(* IEC 61131-3 sources: axsharp/src/AXSharp.compiler/tests/AXSharp.Compiler.CsTests/samples/units/src, 39 files *)

(* ---- compileromitsattribute.st ---- *)
NAMESPACE CompilerOmmits
    {S7.extern=ReadWrite}
    CLASS ClassWithArrays
        VAR PUBLIC
            {#ix-attr:[CompilerOmitsAttribute()]}
            _must_be_omitted_everywhere : Complex;
            {#ix-attr:[CompilerOmitsAttribute("Onliner")]}
            _must_be_omitted_in_onliner : Complex;
            {#ix-attr:[CompilerOmitsAttribute("POCO")]}
             _must_be_omitted_in_poco : Complex;
            _primitive  : ARRAY[0..10] OF BYTE;
        END_VAR

    END_CLASS

    {S7.extern=ReadWrite}
    CLASS PUBLIC Complex
        VAR PUBLIC
            HelloString : STRING;
            Id : ULINT;
        END_VAR
    END_CLASS
END_NAMESPACE

NAMESPACE CompilerOmmitsEnums
    {S7.extern=ReadWrite}
    CLASS ClassWithEnums
        VAR PUBLIC
            colors : Colors;
            NamedValuesColors : NamedValuesColors;
        END_VAR

    END_CLASS

    TYPE
        Colors : (Red, Green, Blue) := Red;
    END_TYPE

    TYPE
        NamedValuesColors : STRING (Red := '1', Green := '2', Blue := '3') := Red;
    END_TYPE

END_NAMESPACE

NAMESPACE CompilerOmmitsMisc
    {S7.extern=ReadWrite}
    CLASS PUBLIC VariousMembers
        VAR PUBLIC
            _SomeClass : SomeClass;
            _Motor : ComersMotor;
        END_VAR
    END_CLASS

    {S7.extern=ReadWrite}
    CLASS SomeClass
        VAR PUBLIC
            SomeClassVariable : STRING;
        END_VAR
    END_CLASS

    TYPE
        {S7.extern=ReadWrite}
        ComersMotor : STRUCT
            isRunning : BOOL;
        END_STRUCT;
        {S7.extern=ReadWrite}
        ComersVehicle : STRUCT
            m : ComersMotor;
            displacement : INT;
        END_STRUCT;
    END_TYPE
END_NAMESPACE

NAMESPACE CompilerOmmitsUnknownArrays
    {S7.extern=ReadWrite}
    CLASS ClassWithArrays
        VAR PUBLIC
            _complexKnown : ARRAY[0..10] OF Complex;
            _complexUnknown : ARRAY [0..10] OF ComplexUnknown;
            _primitive  : ARRAY[0..10] OF BYTE;
        END_VAR

    END_CLASS

    {S7.extern=ReadWrite}
    CLASS PUBLIC Complex
        VAR PUBLIC
            HelloString : STRING;
            Id : ULINT;
        END_VAR
    END_CLASS
END_NAMESPACE

(* ---- enum_simple.st ---- *)
TYPE
    Colors : (Red, Green, Blue) := Red;
END_TYPE

(* ---- misc.st ---- *)
NAMESPACE Enums
{S7.extern=ReadWrite}
    CLASS ClassWithEnums
        VAR PUBLIC
            colors : Colors;
            NamedValuesColors : NamedValuesColors;
        END_VAR

    END_CLASS

    TYPE
        Colors : (Red, Green, Blue) := Red;
    END_TYPE

    TYPE
        NamedValuesColors : STRING (Red := '1', Green := '2', Blue := '3') := Red;
    END_TYPE

END_NAMESPACE

NAMESPACE misc
{S7.extern=ReadWrite}
    CLASS PUBLIC VariousMembers
        VAR PUBLIC
            _SomeClass : SomeClass;
            _Motor : MiscMotor;
        END_VAR
    END_CLASS

    {S7.extern=ReadWrite}
    CLASS SomeClass
        VAR PUBLIC
            SomeClassVariable : STRING;
        END_VAR
    END_CLASS

    TYPE
        {S7.extern=ReadWrite}
        MiscMotor : STRUCT
            isRunning : BOOL;
        END_STRUCT;
        {S7.extern=ReadWrite}
        MiscVehicle : STRUCT
            m : MiscMotor;
            displacement : INT;
        END_STRUCT;
    END_TYPE
END_NAMESPACE

NAMESPACE UnknownArraysShouldNotBeTraspiled
    {S7.extern=ReadWrite}
    CLASS ClassWithArrays
        VAR PUBLIC
            _complexKnown : ARRAY[0..10] OF Complex;
            _complexUnknown : ARRAY [0..10] OF ComplexUnknown;
            _primitive  : ARRAY[0..10] OF BYTE;
        END_VAR

    END_CLASS

    {S7.extern=ReadWrite}
    CLASS PUBLIC Complex
        VAR PUBLIC
            HelloString : STRING;
            Id : ULINT;
        END_VAR
    END_CLASS
END_NAMESPACE

(* ---- mixed_access.st ---- *)
CONFIGURATION config
    VAR_GLOBAL
        {S7.extern=ReadWrite}
        MotorOn : BOOL;             // variable can be read and written

        {S7.extern=ReadOnly}
        MotorState: INT;            // variable can only be read

        MotorFlags: UINT;           // variable is not accessible by an external system (default: hidden)

        {S7.extern=ReadWrite}
        Motor1 : MixedAccessMotor;        // the variables in Motor1 be read and written if enabled

        {S7.extern=ReadOnly}
        Motor2 : MixedAccessMotor;        // the variables in Motor2 be only read if enabled

        {S7.extern=ReadWrite}
        s1 : struct1;
        {S7.extern=ReadWrite}
        s4 : struct4;

        {S7.extern=ReadWrite}
        mot1 : SpecificMotorA;
    END_VAR
END_CONFIGURATION

CLASS MixedAccessMotor
    VAR PUBLIC
        {S7.extern=ReadWrite}
        Run               : BOOL;
        ReverseDirection  : BOOL;
    END_VAR
    VAR INTERNAL
        {S7.extern=ReadOnly}
        ActualVelocity    : LReal;
    END_VAR
    // ...
END_CLASS

TYPE
    struct1 : STRUCT  {S7.extern=ReadWrite}  s2 : struct2;   END_STRUCT;
    struct2 : STRUCT  {S7.extern=ReadOnly}   s3 : struct3;   END_STRUCT;
    struct3 : STRUCT  {S7.extern=ReadWrite}  s4 : struct4;   END_STRUCT;
    struct4 : STRUCT  {S7.extern=ReadWrite}  s5 : INT;       END_STRUCT;
END_TYPE

{S7.extern=ReadWrite}
CLASS ABSTRACT AbstractMotor
    VAR PUBLIC
        Run               : BOOL;
        ReverseDirection  : BOOL;
    END_VAR
    ...
END_CLASS

{S7.extern=ReadWrite}
CLASS GenericMotor  EXTENDS AbstractMotor
    VAR INTERNAL
        {S7.extern=ReadOnly}
        ActualVelocity    : LReal;
    END_VAR
    ...
END_CLASS

{S7.extern=ReadWrite}
CLASS SpecificMotorA  EXTENDS GenericMotor
    VAR INTERNAL
        {S7.extern=ReadWrite}
        MaxAcceleration    : LReal;
    END_VAR
    ...
END_CLASS

(* ---- struct_simple.st ---- *)
TYPE
    {S7.extern=ReadWrite}
    StructSimpleMotor : STRUCT
        isRunning : BOOL;
    END_STRUCT;
    {S7.extern=ReadWrite}
    StructSimpleVehicle : STRUCT
        m : StructSimpleMotor;
        displacement : INT;
    END_STRUCT;
END_TYPE

(* ---- type_named_values.st ---- *)
NAMESPACE NamedValuesNamespace
    TYPE
        LightColors : INT (
            LRED := 12,
            LGREEN := 14,
            LBLUE := 23
        );
    END_TYPE

    {S7.extern=ReadWrite}
    CLASS PUBLIC using_type_named_values
        VAR PUBLIC
            LColors : LightColors;
        END_VAR
    END_CLASS
END_NAMESPACE

(* ---- type_named_values_literals.st ---- *)
NAMESPACE Simatic.Ax.StateFramework
    TYPE
        StateControllerStatus : WORD (
            STATUS_NO_ERR := WORD#16#7000,
            STATUS_IS_RUNNING := WORD#16#7001,
            STATUS_STATE_CHANGED := WORD#16#7002,
            STATUS_NO_INITIALSTATE := WORD#16#8100,
            STATUS_NO_NEXTSTATE := WORD#16#8101
        ) := STATUS_NO_ERR;
    END_TYPE

    {S7.extern=ReadWrite}
    CLASS PUBLIC using_type_named_values
        VAR PUBLIC
            LColors : StateControllerStatus;
        END_VAR
    END_CLASS
END_NAMESPACE

(* ---- type_with_enum.st ---- *)
NAMESPACE Simatic.Ax.StateFramework
    INTERFACE IGuard

        METHOD Check : BOOL
        END_METHOD

        METHOD Reset
        END_METHOD

    END_INTERFACE
END_NAMESPACE

NAMESPACE Simatic.Ax.StateFramework

    /// Condition
    /// GT: Greater than compareValue
    /// EQ: Equal to compareValue
    /// LT: Less than compareValue
    /// NE: Is not equal to compareValue
    /// GE: Greater or equal to compareValue
    /// LE: Less or equal to compareValue
    TYPE
        Condition : (GT, EQ, LT, NE, GE, LE);
    END_TYPE

    {S7.extern=ReadWrite}
    CLASS CompareGuardLint IMPLEMENTS IGuard
        VAR PUBLIC
            Value : REF_TO LINT;
            CompareToValue : LINT;
            Condition : Condition;
        END_VAR

        METHOD PUBLIC Config
            VAR_INPUT
                countValue : REF_TO LINT;
                compareValue : LINT;
                compareCondition : Condition;
            END_VAR
            Value := countValue;
            CompareToValue := compareValue;
            Condition := compareCondition;
        END_METHOD

        // ---------------- IMPLEMENT IGuard---------------------------
        METHOD PUBLIC Check : BOOL

            CASE Condition OF
                Condition#GT : Check := Value^ > CompareToValue;
                Condition#EQ : Check := Value^ = CompareToValue;
                Condition#LT : Check := Value^ < CompareToValue;
                Condition#GE : Check := Value^ >= CompareToValue;
                Condition#LE : Check := Value^ <= CompareToValue;
            END_CASE
            ;

        END_METHOD

        METHOD PUBLIC Reset
            ;
        END_METHOD
        // ---------------- END IMPLEMENT IGuard---------------------------

    END_CLASS
END_NAMESPACE

(* ---- types_with_name_attributes.st ---- *)
NAMESPACE TypeWithNameAttributes
    TYPE
        {#ix-attr:[Container(Layout.Wrap)]}
        {S7.extern=ReadWrite}
        TypesNameAttrMotor : STRUCT
            isRunning : BOOL;
        END_STRUCT;
        {S7.extern=ReadWrite}
        TypesNameAttrVehicle : STRUCT
            m : TypesNameAttrMotor;
            displacement : INT;
        END_STRUCT;
    END_TYPE

    {#ix-prop:public string AttributeName}
    {S7.extern=ReadWrite}
    CLASS NoAccessModifierClass
        VAR PUBLIC
            SomeClassVariable : STRING;
        END_VAR
    END_CLASS
END_NAMESPACE

(* ---- class_extends_and_implements.st ---- *)
{S7.extern=ReadWrite}
CLASS PUBLIC ExtendsAndImplements EXTENDS ExtendeeExtendsAndImplements IMPLEMENTS IImplementation1, IImplementation2

END_CLASS

{S7.extern=ReadWrite}
CLASS PUBLIC ExtendeeExtendsAndImplements

END_CLASS

INTERFACE PUBLIC IImplementation1 END_INTERFACE
INTERFACE PUBLIC IImplementation2 END_INTERFACE

(* ---- class_implements.st ---- *)
{S7.extern=ReadWrite}
CLASS PUBLIC _NULL_CONTEXT IMPLEMENTS IContext

END_CLASS

INTERFACE PUBLIC IContext

END_INTERFACE

(* ---- class_implements_multiple.st ---- *)
{S7.extern=ReadWrite}
CLASS PUBLIC _NULL_CONTEXT_MULTIPLE IMPLEMENTS IContext_Multiple, IObject_Multiple

END_CLASS

INTERFACE PUBLIC IContext_Multiple

END_INTERFACE

INTERFACE PUBLIC IObject_Multiple

END_INTERFACE

(* ---- file_with_unsupported.st ---- *)
NAMESPACE Unsupported
  FUNCTION SomeFunction : INT
    ;
  END_FUNCTION
END_NAMESPACE

(* ---- abstract_members.st ---- *)
{S7.extern=ReadWrite}
CLASS ABSTRACT AbstractMembersMotor
    VAR PUBLIC
        Run               : BOOL;
        ReverseDirection  : BOOL;
    END_VAR
    ...
END_CLASS

(* ---- array_declaration.st ---- *)
NAMESPACE ArrayDeclarationSimpleNamespace
    {S7.extern=ReadWrite}
    CLASS array_declaration_class
        VAR PUBLIC
            primitive : ARRAY[1..100] OF INT;
            complex : ARRAY[1..100] OF some_complex_type;
            // multidimensional arrays should not be transpiled
            complex_multidim : ARRAY[1..100, 0..30] OF some_complex_type;
            primitive_multidim : ARRAY[1..100, 0..100, 0..300] OF INT;
        END_VAR
    END_CLASS
    {S7.extern=ReadWrite}
    CLASS some_complex_type
        VAR

        END_VAR

    END_CLASS

END_NAMESPACE

(* ---- class_all_primitives.st ---- *)
{S7.extern=ReadWrite}
CLASS class_all_primitives
    VAR PUBLIC
        myBOOL	        :       BOOL	      ;
        myBYTE	        :       BYTE	      ;
        myWORD	        :       WORD	      ;
        myDWORD	        :       DWORD	      ;
        myLWORD	        :       LWORD	      ;
        mySINT	        :       SINT	      ;
        myINT	        :       INT	          ;
        myDINT	        :       DINT	      ;
        myLINT	        :       LINT	      ;
        myUSINT	        :       USINT	      ;
        myUINT	        :       UINT	      ;
        myUDINT	        :       UDINT	      ;
        myULINT	        :       ULINT	      ;
        myREAL	        :       REAL	      ;
        myLREAL	        :       LREAL	      ;
        myTIME	        :       TIME	      ;
        myLTIME	        :       LTIME	      ;
        myDATE	        :       DATE	      ;
     //   myLDATE	        :       LDATE	      ;
        myTIME_OF_DAY	:       TIME_OF_DAY	  ;
     //   myLTIME_OF_DAY	:       LTIME_OF_DAY  ;
        myDATE_AND_TIME  :      DATE_AND_TIME ;
     //   myLDATE_AND_TIME :      LDATE_AND_TIME;
     //   myCHAR	        :       CHAR	      ;
     //   myWCHAR	        :       WCHAR	      ;
        mySTRING	        :   STRING	      ;
        myWSTRING	    :       WSTRING	      ;
    END_VAR
END_CLASS

(* ---- class_extended_by_known_type.st ---- *)
USING Simatic.Ax.Stateframework;
USING Simatic.Ax.StatePattern;

NAMESPACE Simatic.Ax.StateFramework
    {S7.extern=ReadWrite}
    CLASS State1Transition EXTENDS AbstractState

        METHOD PUBLIC OVERRIDE OnEntry
            ;
        END_METHOD

        METHOD PUBLIC OVERRIDE OnExit
            ;
        END_METHOD

        METHOD PUBLIC OVERRIDE Action
            ;
        END_METHOD

    END_CLASS

END_NAMESPACE

NAMESPACE Simatic.Ax.StateFramework
    {S7.extern=ReadWrite}
    CLASS ABSTRACT AbstractState IMPLEMENTS IState, IStateMuteable

        VAR PUBLIC
            Transition1 : ITransition;
            StateID : INT;
            StateName : String;
        END_VAR

        VAR PROTECTED
             _actualStatus : StateStatus;
        END_VAR

        // METHOD PUBLIC ABSTRACT OnEntry
        // END_METHOD
        METHOD PUBLIC OnEntry
            _actualStatus := StateStatus#Active;
        END_METHOD

        METHOD PUBLIC ABSTRACT OnExit
        END_METHOD

        METHOD PUBLIC ABSTRACT Action
        END_METHOD

        METHOD PUBLIC GetTransition : ITransition
            VAR_INPUT
                pos : UINT;
            END_VAR
            IF (THIS.TransitionCount() = pos + UINT#1) THEN
                GetTransition := transition1;
            ELSE
                GetTransition := NULL;
            END_IF;
        END_METHOD

        METHOD PUBLIC TransitionCount : UINT
            IF (transition1 <> NULL) THEN
                TransitionCount := UINT#1;
            ELSE
                TransitionCount := UINT#0;
            END_IF;
        END_METHOD

        METHOD PUBLIC GetStateID : INT
            GetStateID := StateID;
        END_METHOD

        METHOD PUBLIC FINAL GetStateName : STRING
            GetStateName := StateName;
        END_METHOD

        METHOD PUBLIC FINAL GetStatus : StateStatus
            GetStatus := _actualStatus;
        END_METHOD

        METHOD PUBLIC FINAL SetStatus
            VAR_INPUT
                status : StateStatus;
            END_VAR
            _actualStatus := status;
        END_METHOD
    END_CLASS
END_NAMESPACE

(* ---- class_extends.st ---- *)
{S7.extern=ReadWrite}
CLASS PUBLIC Extended EXTENDS Extendee

END_CLASS

{S7.extern=ReadWrite}
CLASS PUBLIC Extendee

END_CLASS

(* ---- class_generic_extension.st ---- *)
NAMESPACE Generics
    {#ix-generic:<TOnline, TPlain> where TOnline : ITwinObject}
    {S7.extern=ReadWrite}
    CLASS PUBLIC Extender

    END_CLASS

    {S7.extern=ReadWrite}
    CLASS PUBLIC Extendee EXTENDS Extender
        VAR PUBLIC
            {#ix-generic:TOnline}
            SomeType : SomeType;
            {#ix-generic:TPlain as POCO}
            SomeTypeAsPoco : SomeType;
        END_VAR
    END_CLASS

    {S7.extern=ReadWrite}
    CLASS PUBLIC Extendee2 EXTENDS Extender
        VAR PUBLIC
            {#ix-generic:TOnline}
            {#ix-generic:TPlain as POCO}
            SomeType : SomeType;
        END_VAR
    END_CLASS

    {S7.extern=ReadWrite}
    CLASS SomeType
    END_IF;
END_NAMESPACE

(* ---- class_internal.st ---- *)
{S7.extern=ReadWrite}
CLASS INTERNAL ClassWithComplexTypes

END_CLASS

(* ---- class_no_access_modifier.st ---- *)
{S7.extern=ReadWrite}
CLASS NoAccessModifierClass

END_CLASS

(* ---- class_with_complex_members.st ---- *)
NAMESPACE ClassWithComplexTypesNamespace
    {S7.extern=ReadWrite}
    CLASS PUBLIC ClassWithComplexTypes
        VAR PUBLIC
           myComplexType : ComplexType1;
        END_VAR
    END_CLASS

    {S7.extern=ReadWrite}
    CLASS PUBLIC ComplexType1

    END_CLASS
END_NAMESPACE

(* ---- class_with_constant_members.st ---- *)
NAMESPACE ClassWithConstantMembersNamespace
    {S7.extern=ReadWrite}
    CLASS PUBLIC ClassWithConstantMembers
        VAR PUBLIC
           myNonConstant : INT;
        END_VAR
        VAR CONSTANT
           myConstant : INT := 10;
           myConstantString : STRING := 'hello';
        END_VAR
    END_CLASS
END_NAMESPACE

(* ---- class_with_non_public_members.st ---- *)
NAMESPACE ClassWithNonTraspilableMemberssNamespace
   {S7.extern=ReadWrite}
    CLASS PUBLIC ClassWithNonTraspilableMembers
        VAR PUBLIC
           myComplexType : ComplexType1;
        END_VAR

        VAR
           myComplexType1 : ComplexType1;
           myBooool : BOOL;
        END_VAR

        VAR
           myComplexType2 : ComplexType1;
           myBooool1 : BOOL;
        END_VAR
    END_CLASS
    {S7.extern=ReadWrite}
    CLASS PUBLIC ComplexType1

    END_CLASS
END_NAMESPACE

(* ---- class_with_pragmas.st ---- *)
NAMESPACE ClassWithPragmasNamespace
    {#ix-attr:[Container(Layout.Stack)]}
    {S7.extern=ReadWrite}
    CLASS PUBLIC  ClassWithPragmas
        VAR PUBLIC
           {#ix-attr:[Container(Layout.Wrap)]}
           {S7.extern=ReadWrite}
           myComplexType : ComplexType1;
        END_VAR
    END_CLASS

    CLASS PUBLIC ComplexType1

    END_CLASS
END_NAMESPACE

(* ---- class_with_primitive_members.st ---- *)
NAMESPACE ClassWithPrimitiveTypesNamespace
    {S7.extern=ReadWrite}
    CLASS PUBLIC ClassWithPrimitiveTypes
        VAR PUBLIC
           myBOOL	        :       BOOL	      ;
           myBYTE	        :       BYTE	      ;
           myWORD	        :       WORD	      ;
           myDWORD	        :       DWORD	      ;
           myLWORD	        :       LWORD	      ;
           mySINT	        :       SINT	      ;
           myINT	        :       INT	          ;
           myDINT	        :       DINT	      ;
           myLINT	        :       LINT	      ;
           myUSINT	        :       USINT	      ;
           myUINT	        :       UINT	      ;
           myUDINT	        :       UDINT	      ;
           myULINT	        :       ULINT	      ;
           myREAL	        :       REAL	      ;
           myLREAL	        :       LREAL	      ;
           myTIME	        :       TIME	      ;
           myLTIME	        :       LTIME	      ;
           myDATE	        :       DATE	      ;
           myLDATE	        :       LDATE	      ;
           myTIME_OF_DAY	:       TIME_OF_DAY	  ;
           myLTIME_OF_DAY	:       LTIME_OF_DAY  ;
           myDATE_AND_TIME  :       DATE_AND_TIME ;
           myLDATE_AND_TIME :       LDATE_AND_TIME;
           myCHAR	        :       CHAR	      ;
           myWCHAR	        :       WCHAR	      ;
           mySTRING	        :       STRING	      ;
           myWSTRING	    :       WSTRING	      ;
        END_VAR
    END_CLASS
END_NAMESPACE

(* ---- class_with_using_directives.st ---- *)
{S7.extern=ReadWrite}
CLASS INTERNAL ClassWithUsingDirectives
    USING SimpleFirstLevelNamespace, SimpleQualifiedNamespace.Qualified;
    USING HelloLevelOne.HelloLevelTwo;
    USING InexistingNamespace;
END_CLASS

NAMESPACE SimpleFirstLevelNamespace

END_NAMESPACE

NAMESPACE SimpleQualifiedNamespace.Qualified

END_NAMESPACE

NAMESPACE HelloLevelOne
    NAMESPACE HelloLevelTwo
    END_NAMESPACE
END_NAMESPACE

(* ---- configuration.st ---- *)
CONFIGURATION MyConfiguration
    TASK Main(Interval := T#1000ms, Priority := 1);
    PROGRAM P1 WITH Main: MyProgram;

    VAR_GLOBAL
        {S7.extern=ReadWrite}
        Complex : ComplexForConfig;
        {S7.extern=ReadWrite}
        myBOOL	        :       BOOL	      ;
        {S7.extern=ReadWrite}
        myBYTE	        :       BYTE	      ;
        {S7.extern=ReadWrite}
        myWORD	        :       WORD	      ;
        {S7.extern=ReadWrite}
        myDWORD	        :       DWORD	      ;
        {S7.extern=ReadWrite}
        myLWORD	        :       LWORD	      ;
        {S7.extern=ReadWrite}
        mySINT	        :       SINT	      ;
        {S7.extern=ReadWrite}
        myINT	        :       INT	          ;
        {S7.extern=ReadWrite}
        myDINT	        :       DINT	      ;
        {S7.extern=ReadWrite}
        myLINT	        :       LINT	      ;
        {S7.extern=ReadWrite}
        myUSINT	        :       USINT	      ;
        {S7.extern=ReadWrite}
        myUINT	        :       UINT	      ;
        {S7.extern=ReadWrite}
        myUDINT	        :       UDINT	      ;
        {S7.extern=ReadWrite}
        myULINT	        :       ULINT	      ;
        {S7.extern=ReadWrite}
        myREAL	        :       REAL	      ;
        {S7.extern=ReadWrite}
        myLREAL	        :       LREAL	      ;
        {S7.extern=ReadWrite}
        myTIME	        :       TIME	      ;
        {S7.extern=ReadWrite}
        myLTIME	        :       LTIME	      ;
        {S7.extern=ReadWrite}
        myDATE	        :       DATE	      ;
        {S7.extern=ReadWrite}
        myLDATE	        :       LDATE	      ;
        {S7.extern=ReadWrite}
        myTIME_OF_DAY	:       TIME_OF_DAY	  ;
        {S7.extern=ReadWrite}
        myLTIME_OF_DAY	:       LTIME_OF_DAY  ;
        {S7.extern=ReadWrite}
        myDATE_AND_TIME  :       DATE_AND_TIME ;
        {S7.extern=ReadWrite}
        myLDATE_AND_TIME :       LDATE_AND_TIME;
        {S7.extern=ReadWrite}
        myCHAR	        :       CHAR	      ;
        {S7.extern=ReadWrite}
        myWCHAR	        :       WCHAR	      ;
        {S7.extern=ReadWrite}
        mySTRING	        :       STRING	      ;
        {S7.extern=ReadWrite}
        myWSTRING	    :       WSTRING	      ;
        {S7.extern=ReadWrite}
        mySTRING_10	    :       STRING[10]	  ;
        {S7.extern=ReadWrite}
        myWSTRING_10	:       WSTRING[10]	  ;

        {S7.extern=ReadWrite}
        {#ix-attr:[ReadOnce()]}
        myWSTRING_readOnce	    :       WSTRING	      ;
        {#ix-attr:[ReadOnly()]}
        {S7.extern=ReadWrite}
        myWSTRING_readOnly	    :       WSTRING	      ;
        {#ix-attr:[ReadOnce()]}
        {S7.extern=ReadWrite}
        cReadOnce           : ComplexForConfig;
        {#ix-attr:[ReadOnly()]}
        {S7.extern=ReadWrite}
        cReadOnly           : ComplexForConfig;
        {S7.extern=ReadWrite}
        Colorss : Colorss;
        {S7.extern=ReadWrite}
        Colorsss : Colorsss;

        {S7.extern=ReadWrite}
        {#ix-attr:[CompilerOmitsAttribute()]}
        _must_be_omitted_everywhere : BOOL;
        {S7.extern=ReadWrite}
        {#ix-attr:[CompilerOmitsAttribute("Onliner")]}
        _must_be_omitted_in_onliner : BOOL;
        {S7.extern=ReadWrite}
        {#ix-attr:[CompilerOmitsAttribute("POCO")]}
         _must_be_omitted_in_poco : BOOL;
    END_VAR
END_CONFIGURATION

CONFIGURATION MyConfiguration2
    VAR_GLOBAL
        {S7.extern=ReadWrite}
        Colorss2 : Colorss;
        {S7.extern=ReadWrite}
        Colorsss2 : Colorsss;
    END_VAR
END_CONFIGURATION

{S7.extern=ReadWrite}
CLASS PUBLIC ComplexForConfig
    VAR PUBLIC
        myBOOL	        :       BOOL	      ;
        myBYTE	        :       BYTE	      ;
        myWORD	        :       WORD	      ;
        myDWORD	        :       DWORD	      ;
        myLWORD	        :       LWORD	      ;
        mySINT	        :       SINT	      ;
        myINT	        :       INT	          ;
        myDINT	        :       DINT	      ;
        myLINT	        :       LINT	      ;
        myUSINT	        :       USINT	      ;
        myUINT	        :       UINT	      ;
        myUDINT	        :       UDINT	      ;
        myULINT	        :       ULINT	      ;
        myREAL	        :       REAL	      ;
        myLREAL	        :       LREAL	      ;
        myTIME	        :       TIME	      ;
        myLTIME	        :       LTIME	      ;
        myDATE	        :       DATE	      ;
        myLDATE	        :       LDATE	      ;
        myTIME_OF_DAY	:       TIME_OF_DAY	  ;
        myLTIME_OF_DAY	:       LTIME_OF_DAY  ;
        myDATE_AND_TIME  :       DATE_AND_TIME ;
        myLDATE_AND_TIME :       LDATE_AND_TIME;
        myCHAR	        :       CHAR	      ;
        myWCHAR	        :       WCHAR	      ;
        mySTRING	        :       STRING	      ;
        myWSTRING	    :       WSTRING	      ;
        myMotor         : ConfigMotor;
    END_VAR
END_CLASS

TYPE
    Colorss : (Red, Green, Blue) := Red;
END_TYPE

TYPE
    Colorsss : ULINT (Red := ULINT#1, Green := ULINT#2, Blue := ULINT#3) := Red;
END_TYPE

 TYPE
        {S7.extern=ReadWrite}
        ConfigMotor : STRUCT
            isRunning : BOOL;
        END_STRUCT;
        {S7.extern=ReadWrite}
        ConfigVehicle : STRUCT
            m : ConfigMotor;
            displacement : INT;
        END_STRUCT;
    END_TYPE

(* ---- file_with_usings.st ---- *)
USING FileWithUsingsSimpleFirstLevelNamespace;
USING FileWithUsingsSimpleQualifiedNamespace.Qualified;
USING FileWithUsingsHelloLevelOne.FileWithUsingsHelloLevelTwo;

NAMESPACE FileWithUsingsSimpleFirstLevelNamespace
    CLASS Hello
        VAR

        END_VAR
    END_CLASS
END_NAMESPACE

NAMESPACE FileWithUsingsSimpleQualifiedNamespace.Qualified
    CLASS Hello
        VAR

        END_VAR
    END_CLASS
END_NAMESPACE

NAMESPACE FileWithUsingsHelloLevelOne
    NAMESPACE FileWithUsingsHelloLevelTwo
        CLASS Hello
            VAR

            END_VAR
        END_CLASS
    END_NAMESPACE
END_NAMESPACE

NAMESPACE ExampleNamespace
    CLASS Hello
        VAR
            a : FileWithUsingsSimpleFirstLevelNamespace.Hello;
            b : FileWithUsingsSimpleQualifiedNamespace.Qualified.Hello;
            c : FileWithUsingsHelloLevelOne.FileWithUsingsHelloLevelTwo.Hello;
        END_VAR
    END_CLASS
END_NAMESPACE

(* ---- generics.st ---- *)
// GENERIC
NAMESPACE GenericsTests
    {#ix-generic:<TOnline, TPlain> where TOnline : ITwinObject}
	{S7.extern=ReadWrite}
    CLASS PUBLIC Extender

    END_CLASS

    {S7.extern=ReadWrite}
	CLASS PUBLIC SomeTypeToBeGeneric
	     VAR PUBLIC
		    Boolean : BOOL;
			Cele : INT;
		 END_VAR
	END_CLASS

	{S7.extern=ReadWrite}
   CLASS PUBLIC Extendee2 EXTENDS Extender
        VAR PUBLIC
            {#ix-generic:TOnline}
            {#ix-generic:TPlain as POCO}
            {#ix-attr:[AXOpen.Data.AxoDataEntityAttribute]}
            {#ix-attr:[Container(Layout.Stack)]}
            {#ix-set:AttributeName = "Shared Header"}
            SomeData : SomeTypeToBeGeneric;
        END_VAR
   END_CLASS
END_NAMESPACE

(* ---- makereadonce.st ---- *)
NAMESPACE makereadonce
    {S7.extern=ReadWrite}
    CLASS PUBLIC MembersWithMakeReadOnce
        VAR PUBLIC
            {#ix-attr:[ReadOnce()]}
            makeReadOnceMember : STRING;
            someOtherMember : STRING;

            {#ix-attr:[ReadOnce()]}
            makeReadComplexMember : ComplexMember;
            someotherComplexMember : ComplexMember;
        END_VAR
    END_CLASS
    {S7.extern=ReadWrite}
    CLASS PUBLIC ComplexMember
        VAR PUBLIC
            someMember : STRING;
            someOtherMember : STRING;
        END_VAR
    END_CLASS
END_NAMESPACE

(* ---- makereadonly.st ---- *)
NAMESPACE makereadonly
    {S7.extern=ReadWrite}
    CLASS PUBLIC MembersWithMakeReadOnly
        VAR PUBLIC
            {#ix-attr:[ReadOnly()]}
            makeReadOnceMember : STRING;
            someOtherMember : STRING;

            {#ix-attr:[ReadOnly()]}
            makeReadComplexMember : ComplexMember;
            someotherComplexMember : ComplexMember;
        END_VAR
    END_CLASS
    {S7.extern=ReadWrite}
    CLASS PUBLIC ComplexMember
        VAR PUBLIC
            someMember : STRING;
            someOtherMember : STRING;
        END_VAR
    END_CLASS
END_NAMESPACE

(* ---- multiline_pragmas.st ---- *)
// GENERIC
NAMESPACE MultilinePragmas
   {S7.extern=ReadWrite}
   CLASS PUBLIC Extendee2 EXTENDS Extender
        VAR PUBLIC
            {#ix-set:PlcTextList = "[1]:'<#Messenger 1: message text for message code 1#>':'<#Messenger 1: help text for message code 1#>';
                                    [2]:'<#Messenger 1: message text for message code 2#>':'<#Messenger 1: help text for message code 2#>';
                                    [3]:'<#Messenger 1: message text for message code 3#>':'<#Messenger 1: help text for message code 3#>';
                                    [4]:'<#Messenger 1: message text for message code 4#>':'<#Messenger 1: help text for message code 4#>';
                                    [5]:'<#Messenger 1: message text for message code 5#>':'<#Messenger 1: help text for message code 5#>';
                                    [6]:'<#Messenger 1: message text for message code 6#>':'<#Messenger 1: help text for message code 6#>';
                                    [7]:'<#Messenger 1: message text for message code 7#>':'<#Messenger 1: help text for message code 7#>';
                                    [8]:'<#Messenger 1: message text for message code 8#>':'<#Messenger 1: help text for message code 8#>';
                                    [9]:'<#Messenger 1: message text for message code 9#>':'<#Messenger 1: help text for message code 9#>';
                                    [10]:'<#Messenger 1: message text for message code 10#>':'<#Messenger 1: help text for message code 10#>';
                                    [11]:'<#Messenger 1: message text for message code 11#>':'<#Messenger 1: help text for message code 11#>'"}
            _messge : INT;
        END_VAR
   END_CLASS
END_NAMESPACE

(* ---- ref_to_simple.st ---- *)
NAMESPACE RefToSimple
    {S7.extern=ReadWrite}
    CLASS ref_to_simple
        VAR PUBLIC
            a : REF_TO INT;
            b : REF_TO referenced;
        END_VAR
    END_CLASS

    {S7.extern=ReadWrite}
    CLASS referenced
        VAR PUBLIC
            b : INT;
        END_VAR
    END_CLASS
END_NAMESPACE

(* ---- simple_empty_class.st ---- *)
{S7.extern=ReadWrite}
CLASS PUBLIC simple_class
END_CLASS

(* ---- simple_empty_class_within_namespace.st ---- *)
NAMESPACE sampleNamespace
    {S7.extern=ReadWrite}
    CLASS PUBLIC simple_empty_class_within_namespace
    END_CLASS
END_NAMESPACE

(* ---- string_capacity.st ---- *)
NAMESPACE StringCapacityNamespace
    {S7.extern=ReadWrite}
    CLASS PUBLIC ClassWithDeclaredStringCapacities
        VAR PUBLIC
            myString10      :   STRING[10];
            myWString10     :   WSTRING[10];
            myString        :   STRING;
            myWString       :   WSTRING;
            myWString1000   :   WSTRING[1000];
            myString10Array :   ARRAY[0..3] OF STRING[10];
        END_VAR
    END_CLASS
END_NAMESPACE

(* ---- types_with_property_attributes.st ---- *)
NAMESPACE TypesWithPropertyAttributes
    {#ix-prop:public string Description}
    {#ix-set:Description = "Some added property name value"}
    {S7.extern=ReadWrite}
    CLASS SomeAddedProperties
        VAR PUBLIC
            {#ix-set:AttributeName = "Pocitadlo"}
            Counter : INT;
        END_VAR
    END_CLASS
END_NAMESPACE

(* ---- program.st ---- *)
PROGRAM MyProgram
    VAR_EXTERNAL

    END_VAR

    VAR

    END_VAR

    VAR_TEMP

    END_VAR

    // code here
    ;
END_PROGRAM
